TYPE ST_ConvPersist :
STRUCT
	// Nastawy operatora
	Cfg		: ST_ConvCfg;

	// Pamiec stanu maszyny
	Mem		: ST_ConvMem;
END_STRUCT
END_TYPE

(* stored: Version 1.1.0.1
   DUT ST_ConvPersist: Id {7a1c0007-0000-4000-9000-000000000007} *)
